(* IEC 61131-3 sources: axsharp/src/AXSharp.compiler/tests/AXSharp.CompilerTests/samples/plt/lib/src, 1 file *)

(* ---- library.st ---- *)
NAMESPACE MyLibrary

    CLASS PUBLIC MyClass
        VAR PUBLIC

        END_VAR

        VAR PRIVATE

        END_VAR

        METHOD PUBLIC MyMethod : BOOL
            MyMethod := FALSE;
        END_METHOD
    END_CLASS

END_NAMESPACE
